// TIA Portal V17 export
// export: Created 2026-11-17T10:42:02.8543703Z, ExportSetting WithDefaults, DisplayName Totally Integrated Automation Portal, DisplayVersion V17, DisplayName TIA Portal Openness, DisplayVersion V17, DisplayName TIA Portal Version Control Interface, DisplayVersion V17, DisplayName STEP 7 Professional, DisplayVersion V17, DisplayName STEP 7 Safety, DisplayVersion V17, DisplayName WinCC Advanced, DisplayVersion V17
VAR_GLOBAL   // PLC tag table "红绿灯变量表"
   StartPB AT %M0.0 : Bool;   // HMI 启动按钮
   StopPB AT %M0.1 : Bool;   // HMI 停止按钮
   Run AT %M0.2 : Bool;   // 运行自锁与指示灯
   NS_Red AT %Q0.0 : Bool;   // 南北红灯
   NS_Yellow AT %Q0.1 : Bool;   // 南北黄灯
   NS_Green AT %Q0.2 : Bool;   // 南北绿灯
   EW_Red AT %Q0.3 : Bool;   // 东西红灯
   EW_Yellow AT %Q0.4 : Bool;   // 东西黄灯
   EW_Green AT %Q0.5 : Bool;   // 东西绿灯
   Done1 AT %M1.0 : Bool;   // 东西绿灯定时到
   Done2 AT %M1.1 : Bool;   // 东西黄灯定时到
   Done3 AT %M1.2 : Bool;   // 南北绿灯定时到
   Done4 AT %M1.3 : Bool;   // 南北黄灯定时到
END_VAR
